Staubli VAL3: start.pgx

public program start()
  local string l_sArmType
  local string l_sSeries
begin
  //****************************************************************************************
  // +-----------------------------------------------------------------------------------+
  // !                                 Stäubli SmartTCP                                  !
  // !                                                                                   !
  // !                Copyright by  Stäubli(Hagnzhou) Mechatronic Co.,Ltd.               !
  // +-----------------------------------------------------------------------------------+
  // General description：  Stäubli TCP calibration application for TX2/TS2 robot
  // Developer:             ZhangHuaJun
  // Application version：  V1.2
  // Application Date:      February 24, 2020
  // Hardware required：    TX2/TS2-CS9-SP2 Robot
  // Software required：    Val3 s8.8.3+
  // VAL3 Addons：          Expansion
  // Fieldbus required:     None
  // VAL3 Options：         None
  // Included libraries：   None
  // Miscellaneous：        None
  //****************************************************************************************
  l_sArmType=getVersion("Arm Type")
  if l_sArmType!=""
    l_sSeries=left(l_sArmType,3)
    switch l_sSeries
      case "ts2"
        call ts2:start()
      break
      case "tx2"
        call tx2:start()
      break
    endSwitch
  endIf
end
